// TIA Portal V21 export
Screen "T10_RectV"  1024x768, Number=30
  ScreenLayer 
    Rectangle "P_CraneY" at 0,0 size 100x30
      VerticalMovementAnimation   RangeTo=9, Tag=CraneY
